Fanuc KAREL source: kt00903.KL

PROGRAM KT00903
%STACKSIZE=65535
%PRIORITY=65535
%NOLOCKGROUP
VAR
P1 : POSITION
P2 : POSITION
OUT : VECTOR
BEGIN
OUT=APPROACH(P1)
END KT00903
